Fanuc KAREL source: kf00080.KL

-- PROVISIONAL review KL for V1013-1; original PC SHA256 cf751d4f8e52dd3f21211c3ab139c8f4072e09d94014559460bcc60ccf528fb8
-- Incomplete behavior may be omitted. Consult companion uncertainty JSON. Do not deploy.
PROGRAM KF00080
%NOLOCKGROUP
BEGIN
  -- UNRESOLVED_PC offsets 5-15; opcodes 27,22,31
  -- UNRESOLVED_PC offsets 20-24; opcodes 7F
END KF00080
